PROGRAM TESTS_MAIN
VAR
{IF defined (Tests)}
	startTests : BOOL;
	// FBs to test
	fbMovingAverageTest 					: FB_MovingAverage_Test;
	fbConsumptionCalculatorTest 			: FB_ConsumptionCalculator_Test;
	fbmFTest 								: FB_mF_Test;
	fbCo2ModelDeviationHandlerTest 			: FB_Co2FlowModelDeviationHandler_Test;
	fbAutomaticExtractionStateMachineTest 	: FB_AutomaticExtractionStateMachine_Test;
	fbRuntimeTest 							: FB_Runtime_Test;
	fbControlValveStateMachineTest			: FB_ControlValveStateMachine_Test;
	fbReactorValvesTest						: FB_ReactorValves_Test;
	
	// Handlers to test
	AutomaticExtractionHandlerTest			: AutomaticExtractionHandler_Test;
	
	movingavg 						: FB_MovingAverage;
	consumptioncalc 				: FB_ConsumptionCalculator;
	measF : REAL;
	mF : FB_mF;
	TON_Test : TON;
	meas : LREAL;
	uTest : ARRAY[1..15] OF LREAL;
	fbGetCurTaskIndex : GETCURTASKINDEX;
{END_IF}
END_VAR


fbGetCurTaskIndex();
IF _TaskInfo[fbGetCurTaskIndex.index].FirstCycle THEN
    // The code that you want to be executed at the first cycle
	mF.setParams(
		activateObserver := FALSE);
END_IF

IF startTests THEN
	TcUnit.RUN();
	movingavg.startCalculation(
							start := TRUE,
							measurement := meas,
							intervalS := 1,
							windowS := 10,
							dTime := T#10MS,
							excludeUntilReady := FALSE);
	consumptioncalc.calculate(
							start := TRUE,
							valuePerSec := movingavg.value/60,
							intervalS := 10,
							dtime := T#10MS);
	uTest[1];
	TON_Test(IN := TRUE, PT := T#1S);
	IF TON_Test.Q THEN
		mF.Step(
				u := uTest,
				yMeas := meas);
		TON_Test(IN := FALSE);
		mF.y[1];
	END_IF
END_IF

END_PROGRAM

(* stored: Version 1.1.0.1, ProductVersion 3.1.4024.9
   POU TESTS_MAIN: Id {c34b9cd4-20c9-4aab-a9d3-84efa1ac7435}, SpecialFunc None *)
